Fanuc KAREL source: kt00001.KL

-- PROVISIONAL review KL for V1013-1; original PC SHA256 bc56e5cccf98dcfdda539ee1205a5655163817f752445b292aece96278ae6268
-- Incomplete behavior may be omitted. Consult companion uncertainty JSON. Do not deploy.
PROGRAM KT00001
%NOLOCKGROUP
VAR
  I1 : INTEGER
  I2 : INTEGER
  OUT : INTEGER
BEGIN
  -- UNRESOLVED_PC offsets 5-16; opcodes 2E,23
  -- UNRESOLVED_PC offsets 21-32; opcodes 2E,23
  -- UNRESOLVED_PC offsets 37-48; opcodes 2E,23
  -- UNRESOLVED_PC offsets 53-64; opcodes 2E,23
  -- UNRESOLVED_PC offsets 69-88; opcodes 21,21,52,23
  -- UNRESOLVED_PC offsets 93-97; opcodes 7F
END KT00001
